// Mitsubishi GX Works2 project: 20261012_기초회로_인터록 회로_선입우선   PLC: Q03UDV

PROGRAM MAIN
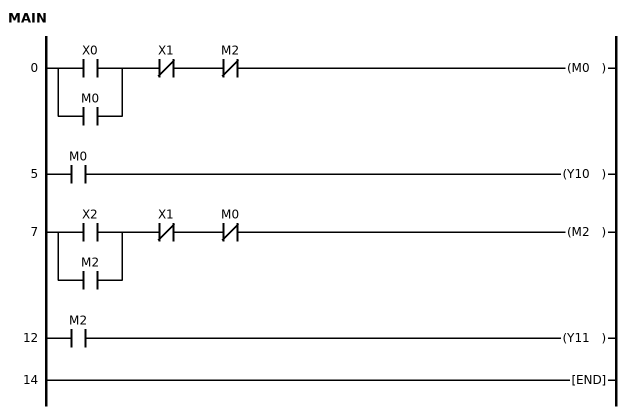
0     LD      X0
      OR      M0
      ANI     X1
      ANI     M2
      OUT     M0
5     LD      M0
      OUT     Y10
7     LD      X2
      OR      M2
      ANI     X1
      ANI     M0
      OUT     M2
12    LD      M2
      OUT     Y11
14    END
END_PROGRAM
